Fanuc KAREL source: KT00143.KL

PROGRAM KT00143
%NOLOCKGROUP
VAR
  R1: REAL
  H2: ARRAY[2] OF SHORT
  OUT: INTEGER
BEGIN
  R1 = 2.0
    H2[1] = 3
  OUT = R1 DIV H2[1]
END KT00143
